Fanuc KAREL source: KT00734.KL

PROGRAM KT00734
%NOLOCKGROUP
VAR
  ARG: ARRAY[4] OF BOOLEAN
  OUT: BOOLEAN
BEGIN
  OUT = UNINIT(ARG)
END KT00734
